Staubli VAL3: cycle_End.pgx

program cycle_End()
begin

  //cycle进程:Ending
  rs:_nOmacStat=7
  _bEndCycle=true
  wait(taskStatus("Main")<0)

  // Stop task
  stopMove()
  call ar:getCurMoveID(bGetMovId,"End")
  wait(isSettled())
  resetMotion()
  //shutdown arm power
  disablePower()

  //cycle进程:Stopped
  rs:_nOmacStat=9
  logMsg("当前处于停止状态 "+toString(".2",clock()))
  rs:_sRobotStatus="当前处于停止状态"
end
